(* IEC 61131-3 sources: IRIS-Project/LASAL CONTROL SOFTWARE/LasalProject_2025_09_25/Network, 1 file *)

(* ---- ConfigObjects.st ---- *)
FUNCTION GLOBAL TAB TASK_CONF
_K_TASK, _K_REAL,
_K_END_VAR,

_K_TASK, _K_CYCLIC,
_K_END_VAR,

_K_TASK, _K_BACKGROUND,
_K_END_VAR,

_K_END_CONF
END_FUNCTION

FUNCTION GLOBAL TAB IPR_CONF
_K_IPR
	0$UINT,
_K_END_VAR,
_K_END_CONF
END_FUNCTION

FUNCTION GLOBAL TAB CONFIG_TABLES
00114$UINT,
0$UINT, 1, 58, "_AXISBASE",
0$UINT, 0, 4, "_CAN",
0$UINT, 1, 10, "_CANLIB",
0$UINT, 1, 0, "_CHECKSUM",
0$UINT, 1, 20, "_FILESYS",
0$UINT, 0, 5, "_LINKER",
0$UINT, 1, 0, "_LMCABSENCODER",
0$UINT, 1, 114, "_LMCAXIS",
0$UINT, 2, 105, "_LMCAXISBASE",
0$UINT, 1, 32, "_LMCAXISREF",
0$UINT, 1, 40, "_LMCAXISVIS",
0$UINT, 1, 62, "_LMCAXISVISINT",
0$UINT, 1, 0, "_LMCAXISVISLOGHANDLE",
0$UINT, 1, 0, "_LMCAXISVISLOGVIEWER",
0$UINT, 1, 13, "_LMCAXISVISPARA",
0$UINT, 1, 1, "_LMCAXISVOVMONITORING",
0$UINT, 1, 75, "_LMCMATHFUNCTIONS",
0$UINT, 1, 0, "_LMCMODULEBASE",
0$UINT, 1, 0, "_LMCPUBLISHER",
0$UINT, 1, 11, "_LMCREFBASE",
0$UINT, 1, 21, "_LMCSAFETY",
0$UINT, 1, 36, "_MODBUSTCPSLAVE",
0$UINT, 1, 1, "_MULTITASK",
0$UINT, 0, 5, "_OSKERNEL",
0$UINT, 1, 34, "_SERLIB",
0$UINT, 0, 0, "_STDLIB",
0$UINT, 0, 0, "_SYSMSG",
0$UINT, 1, 1, "_TASKOBJECTCONTROL",
0$UINT, 1, 38, "_TCPIP_SERVER",
0$UINT, 1, 18, "AI084",
0$UINT, 1, 21, "ASCII_BIN",
0$UINT, 0, 0, "ATTUATORE",
0$UINT, 0, 0, "AUTOMANSELECTOR",
0$UINT, 0, 0, "AUTOMATIC_STEP_SETTINGS",
0$UINT, 2, 1, "BUSINTERFACESDIASINTERNAL",
0$UINT, 1, 46, "CONTROLLER",
0$UINT, 0, 0, "CONTROLLOSERVERMODBUS",
0$UINT, 1, 1, "CP112_IOS",
0$UINT, 0, 4, "CRITICALSECTION",
0$UINT, 1, 12, "DI160",
0$UINT, 2, 33, "DIASMASTER",
0$UINT, 1, 83, "DIASMASTERC",
0$UINT, 2, 25, "DIASMASTERMAIN",
0$UINT, 1, 0, "DIASMASTERPOSTSCAN",
0$UINT, 0, 0, "DISCHARGETIMER",
0$UINT, 1, 11, "EEPROM",
0$UINT, 0, 0, "ESTOPMANAGER",
0$UINT, 0, 0, "EXACTSTEP",
0$UINT, 0, 0, "HOLDINGREGISTER",
0$UINT, 0, 0, "HOLDINGREGISTER_2",
0$UINT, 0, 0, "HOLDINGREGISTER_3",
0$UINT, 1, 21, "HUB_BASE",
0$UINT, 2, 11, "HUB_BASE_ROOT",
0$UINT, 2, 36, "HWBASE",
0$UINT, 2, 56, "HWBASECDIAS",
0$UINT, 1, 0, "HWCLOGGING",
0$UINT, 5, 21, "HWCONTROL",
0$UINT, 1, 10, "HWCONTROLBASE",
0$UINT, 1, 0, "HWRTPOSTSCAN",
0$UINT, 1, 6, "I2CCDIAS",
0$UINT, 0, 0, "INPUTREGISTER",
0$UINT, 0, 0, "IRRADIATIONMANAGER",
0$UINT, 1, 0, "LOGIC_NOT",
0$UINT, 1, 0, "LOGIC_XOR",
0$UINT, 0, 0, "MAINSEQUENCE",
0$UINT, 0, 0, "MANAGER_GLOBALE",
0$UINT, 0, 0, "MANAGER_MANUAL_MOTOR",
0$UINT, 0, 0, "MANAGERMOTORI",
0$UINT, 0, 0, "MANUAL_MOTOR",
0$UINT, 0, 0, "MANUAL_MOTORBT",
0$UINT, 0, 0, "MANUAL_STEP_SETTINGS",
0$UINT, 0, 0, "MANUALMOTOR_CBCM",
0$UINT, 0, 0, "MANUALMOTOR_DB",
0$UINT, 1, 22, "MERKEREX",
0$UINT, 0, 0, "MODE_SELECTOR_CLASS",
0$UINT, 0, 0, "MOTORE_M1",
0$UINT, 0, 0, "MOTORE_M2",
0$UINT, 0, 0, "MOTORE_M3",
0$UINT, 0, 0, "MOTORE_M4",
0$UINT, 0, 0, "MOTORE_M5",
0$UINT, 0, 0, "MOTORE_M6",
0$UINT, 0, 0, "MOTORE_M7",
0$UINT, 0, 0, "MOVETIMER",
0$UINT, 0, 0, "MPS",
0$UINT, 0, 0, "RACK12V",
0$UINT, 1, 9, "RAMFILE",
0$UINT, 0, 0, "RESET",
0$UINT, 3, 19, "SAFETYCDIAS_BASE",
0$UINT, 2, 26, "SAFETYMANAGER",
0$UINT, 1, 4, "SAFETYUDP",
0$UINT, 1, 60, "SDIASBASE",
0$UINT, 1, 10, "SDIASHUBBASE",
0$UINT, 1, 97, "SDIASMANAGER",
0$UINT, 2, 6, "SDIASPLC",
0$UINT, 0, 42, "SIGCLIB",
0$UINT, 1, 6, "ST151",
0$UINT, 1, 0, "ST151_INTVISU",
0$UINT, 1, 4, "ST151BASE",
0$UINT, 1, 3, "STEPPERCONTROL",
0$UINT, 1, 11, "STRING",
0$UINT, 1, 85, "STRINGINTERNAL",
0$UINT, 1, 21, "SYNCCALL",
0$UINT, 1, 5, "SYSDATETIME",
0$UINT, 0, 1, "SYSTEM",
0$UINT, 1, 1, "TIMEDATELIB",
0$UINT, 1, 0, "TIMERLIB",
0$UINT, 1, 44, "TO127",
0$UINT, 2, 20, "VARAN_BASE",
0$UINT, 3, 7, "VARANMANAGER",
0$UINT, 2, 7, "VARANMANAGER_1",
0$UINT, 1, 26, "VARANMANAGER_BASE",
0$UINT, 1, 3, "VIRTUALBASEINIT",
0$UINT, 2, 11, "WATCHDOGDIAS",
0$UINT, 1, 1, "XXXBASE_IOS",
ONE_CFG$UINT, 0, 0, "ONE_Comunicazione_ModBus",
ONE_CFG$UINT, 0, 0, "ONE_HW_Network",
ONE_CFG$UINT, 0, 0, "ONE_IRIS_MANAGER",
ONE_CFG$UINT, 0, 0, "ONE_Manual",
ONE_CFG$UINT, 0, 0, "ONE_Profili_Assi",
ONE_CFG$UINT, 0, 0, "ONE_Settings",
ONE_CFG$UINT, 0, 0, "ONE_Timer",
TASK_CFG$UINT, 0, 0, "TASK_CONF",
IPR_CFG$UINT, 0, 0, "IPR_CONF",
PRJ_CFG$UINT, 0, 0, "v1",
END_FUNCTION

#ifdef __LSLLDR_IOELEMENTS__
FUNCTION GLOBAL TAB _IO_ELEMENTS_TAB
0001$UINT, 0133$UINT,
"**IOCONN_EMPTY**", "ST1517.Input1",
"IO_Element", "_LMCAxis_M1.Control",
"IO_Element0", "ST1511.AxError",
"IO_Element1", "ST1511.Enable",
"IO_Element10", "_LMCAxis_M7.Control",
"IO_Element100", "_LMCAxis_M6.ActPos",
"IO_Element101", "Manager_globale1.enable",
"IO_Element102", "_LMCAxis_M1.ActPos",
"IO_Element103", "_LMCAxis_M2.ActPos",
"IO_Element104", "_LMCAxis_M3.ActPos",
"IO_Element105", "_LMCAxis_M4.ActPos",
"IO_Element106", "_LMCAxis_M5.ActPos",
"IO_Element107", "_LMCAxis_M6.ActPos",
"IO_Element108", "_LMCAxis_M7.ActPos",
"IO_Element109", "TO1271.Output4",
"IO_Element11", "ST1511.ActPosition",
"IO_Element110", "TO1271.Output8",
"IO_Element111", "TO1271.Output11",
"IO_Element112", "TO1271.Output10",
"IO_Element113", "ST1516.MaxCurrent",
"IO_Element114", "MPS1.ReqToMPS",
"IO_Element115", "Motore_M51.s_TabletTimer",
"IO_Element116", "Manager_globale1.ComandoIrradiation",
"IO_Element117", "MoveTimer1.s_StartStopTimer",
"IO_Element118", "MoveTimer1.s_StartStopTimer",
"IO_Element119", "MainSequence1.s_EasyGUI",
"IO_Element12", "_LMCAxis_M1.Control",
"IO_Element120", "IrradiationTimers.s_EasyGUI",
"IO_Element121", "Reset1.s_ResetT",
"IO_Element122", "IrradiationTimers.s_TimerStartStop",
"IO_Element123", "ST1514.MaxCurrent",
"IO_Element124", "ST1511.MaxCurrent",
"IO_Element125", "ST1513.MaxCurrent",
"IO_Element126", "ST1516.MaxCurrent",
"IO_Element127", "ST1515.MaxCurrent",
"IO_Element128", "ST1512.MaxCurrent",
"IO_Element129", "MoveTimer1.s_1_3_pelletMode",
"IO_Element13", "ST1511.Input2",
"IO_Element130", "IrradiationTimers.s_1_3_pelletMode",
"IO_Element14", "Motore_M11.M1_Correction_Step",
"IO_Element15", "ST1512.ActPosition",
"IO_Element16", "ST1511.Input1",
"IO_Element17", "ST1511.Input2",
"IO_Element18", "Motore_M41.M4_Correction_Step",
"IO_Element19", "DI1601.Input3",
"IO_Element2", "ST1511.SetFreqOut",
"IO_Element20", "ST1512.AxError",
"IO_Element21", "ST1512.Enable",
"IO_Element22", "ST1512.SetFreqOut",
"IO_Element23", "ST1512.ErrorQuit",
"IO_Element24", "ST1513.ActPosition",
"IO_Element25", "ST1513.AxError",
"IO_Element26", "ST1513.Enable",
"IO_Element27", "ST1513.SetFreqOut",
"IO_Element28", "ST1513.ErrorQuit",
"IO_Element29", "ST1514.ActPosition",
"IO_Element3", "ST1511.ErrorQuit",
"IO_Element30", "ST1514.AxError",
"IO_Element31", "ST1514.Enable",
"IO_Element32", "ST1514.SetFreqOut",
"IO_Element33", "ST1514.ErrorQuit",
"IO_Element34", "ST1512.Input2",
"IO_Element35", "TO1271.Output2",
"IO_Element36", "ST1513.Input1",
"IO_Element37", "ST1513.Input2",
"IO_Element38", "ST1514.Input1",
"IO_Element39", "TO1271.Output3",
"IO_Element4", "_LMCAxis_M2.Control",
"IO_Element40", "TO1271.Output1",
"IO_Element41", "TO1271.Output5",
"IO_Element42", "TO1271.Output6",
"IO_Element43", "TO1271.Output7",
"IO_Element44", "ST1515.ActPosition",
"IO_Element45", "ST1515.AxError",
"IO_Element46", "ST1515.Enable",
"IO_Element47", "ST1515.SetFreqOut",
"IO_Element48", "ST1515.ErrorQuit",
"IO_Element49", "ST1515.Input1",
"IO_Element5", "_LMCAxis_M3.Control",
"IO_Element50", "ST1516.Input1",
"IO_Element51", "ST1516.Input2",
"IO_Element52", "ST1513.MaxCurrent",
"IO_Element53", "ST1516.ActPosition",
"IO_Element54", "ST1516.AxError",
"IO_Element55", "ST1516.Enable",
"IO_Element56", "ST1516.SetFreqOut",
"IO_Element57", "ST1516.ErrorQuit",
"IO_Element58", "ST1511.MaxCurrent",
"IO_Element59", "ST1515.MaxCurrent",
"IO_Element6", "_LMCAxis_M4.Control",
"IO_Element60", "_LMCAxis_M5.ActPos",
"IO_Element61", "_LMCAxis_M1.ActPos",
"IO_Element62", "_LMCAxis_M3.ActPos",
"IO_Element63", "ST1517.ActPosition",
"IO_Element64", "ST1517.AxError",
"IO_Element65", "ST1517.Enable",
"IO_Element66", "ST1517.SetFreqOut",
"IO_Element67", "ST1517.ErrorQuit",
"IO_Element68", "ST1517.Input1",
"IO_Element69", "ST1517.Input2",
"IO_Element7", "_LMCAxis_M5.Control",
"IO_Element70", "_LMCAxis_M7.ActPos",
"IO_Element71", "ST1514.MaxCurrent",
"IO_Element72", "Motore_M31.M3_Correction_Step",
"IO_Element73", "Motore_M51.M5_ChargingCorrection_step_1",
"IO_Element74", "Motore_M51.M5_ChargingCorrection_step_2",
"IO_Element75", "Motore_M51.M5_ChargingCorrection_step_3",
"IO_Element76", "Motore_M51.M5_IrradiationCorrection_step_1",
"IO_Element77", "Motore_M51.M5_IrradiationCorrection_step_2",
"IO_Element78", "_LMCAxis_M2.Control",
"IO_Element79", "Motore_M51.M5_IrradiationCorrection_step_3",
"IO_Element8", "_LMCAxis_M6.Control",
"IO_Element80", "Motore_M51.M5_DischargeCorrection_step",
"IO_Element81", "ST1512.Input2",
"IO_Element82", "_LMCAxis_M3.Control",
"IO_Element83", "_LMCAxis_M4.Control",
"IO_Element84", "DI1601.Input1",
"IO_Element85", "TO1271.Output9",
"IO_Element86", "_LMCAxis_M5.Control",
"IO_Element87", "_LMCAxis_M6.Control",
"IO_Element88", "_LMCAxis_M7.Control",
"IO_Element89", "ST1513.Input1",
"IO_Element9", "ST1511.Input1",
"IO_Element90", "ST1513.Input2",
"IO_Element91", "ST1514.Input1",
"IO_Element92", "ST1515.Input1",
"IO_Element93", "ST1516.Input1",
"IO_Element94", "ST1516.Input2",
"IO_Element95", "Motore_M51.s_tablet_irradiation_position",
"IO_Element96", "DischargeTimer1.s_StartStopTimer",
"IO_Element97", "_LMCAxis_M2.ActPos",
"IO_Element98", "ManagerMotori1.From_MPS",
"IO_Element99", "_LMCAxis_M4.ActPos",
0134$UINT,
"**IOCONN_EMPTY**", "M7_Target_Block.M_LS_1",
"**IOCONN_EMPTY**", "M7_Target_Block.M_LS_2",
"IO_Element", "Motore_M11.Comando_M1",
"IO_Element0", "StepperControl_M1.HWErrors",
"IO_Element1", "StepperControl_M1.Active",
"IO_Element10", "Motore_M71.Comando_M7",
"IO_Element100", "Motore_M61.SetPosition_Controller",
"IO_Element101", "AutoManSelector1.toAutomatic",
"IO_Element102", "M1_Charge_Slider.setPositionController",
"IO_Element103", "M2_Charge_Buffer.setPositionController",
"IO_Element104", "M3_Discharge_Slider.setPositionController",
"IO_Element105", "M4_Discharge_Buffer.setPositionController",
"IO_Element106", "M5_Central_Movement.setPositionController",
"IO_Element107", "M6_Longitudinal_axis.setPositionController",
"IO_Element108", "M7_Target_Block.setPositionController",
"IO_Element109", "Rack12V1.ToPLC",
"IO_Element11", "_LMCAxis_M1.ActPosition",
"IO_Element110", "ManagerMotori1.LED_Rosso",
"IO_Element111", "ManagerMotori1.LED_Arancione",
"IO_Element112", "ManagerMotori1.LED_Verde",
"IO_Element113", "MPS1.To_CameraAlignment_Power",
"IO_Element114", "ManagerMotori1.c_MPS_Req",
"IO_Element115", "IrradiationTimers.NrIrrTablets",
"IO_Element116", "IrradiationTimers.SetStartStopIrr",
"IO_Element117", "Motore_M51.c_TimerMov",
"IO_Element118", "Motore_M41.c_TimerMov",
"IO_Element119", "AutoManSelector1.c_EasyGUIEn_MainS",
"IO_Element12", "M1_Charge_Slider.Comando_Motore",
"IO_Element120", "AutoManSelector1.c_EasyGUIEn_IrrT",
"IO_Element121", "Manager_globale1.c_ResetTimer",
"IO_Element122", "Motore_M51.c_TimerIrr",
"IO_Element123", "M4_Discharge_Buffer.c_MaxCurrent",
"IO_Element124", "M1_Charge_Slider.c_MaxCurrent",
"IO_Element125", "M3_Discharge_Slider.c_MaxCurrent",
"IO_Element126", "M6_Longitudinal_axis.c_MaxCurrent",
"IO_Element127", "M5_Central_Movement.c_MaxCurrent",
"IO_Element128", "M2_Charge_Buffer.c_MaxCurrent",
"IO_Element129", "ManagerMotori1.c_1_3_pelletMode_TimerMov",
"IO_Element13", "Motore_M11.M1_LS_2",
"IO_Element130", "ManagerMotori1.c_1_3_pelletMode_TimerIrr",
"IO_Element14", "Automatic_Step_Settings1.c_M1_Correction_Step",
"IO_Element15", "_LMCAxis_M2.ActPosition",
"IO_Element16", "M1_Charge_Slider.M_LS_1",
"IO_Element17", "M1_Charge_Slider.M_LS_2",
"IO_Element18", "Automatic_Step_Settings1.c_M4_Correction_Step",
"IO_Element19", "Manager_globale1.Reset_IN",
"IO_Element2", "StepperControl_M1.OutputSignal",
"IO_Element20", "StepperControl_M2.HWErrors",
"IO_Element21", "StepperControl_M2.Active",
"IO_Element22", "StepperControl_M2.OutputSignal",
"IO_Element23", "StepperControl_M2.HWErrorQuit",
"IO_Element24", "_LMCAxis_M3.ActPosition",
"IO_Element25", "StepperControl_M3.HWErrors",
"IO_Element26", "StepperControl_M3.Active",
"IO_Element27", "StepperControl_M3.OutputSignal",
"IO_Element28", "StepperControl_M3.HWErrorQuit",
"IO_Element29", "_LMCAxis_M4.ActPosition",
"IO_Element3", "StepperControl_M1.HWErrorQuit",
"IO_Element30", "StepperControl_M4.HWErrors",
"IO_Element31", "StepperControl_M4.Active",
"IO_Element32", "StepperControl_M4.OutputSignal",
"IO_Element33", "StepperControl_M4.HWErrorQuit",
"IO_Element34", "Motore_M21.M2_LS",
"IO_Element35", "Attuatore1.R_aus_1",
"IO_Element36", "Motore_M31.M3_LS_1",
"IO_Element37", "Motore_M31.M3_LS_2",
"IO_Element38", "Motore_M41.M4_LS",
"IO_Element39", "Attuatore1.R_aus_2",
"IO_Element4", "Motore_M21.Comando_M2",
"IO_Element40", "Attuatore1.R_p",
"IO_Element41", "Attuatore2.R_p",
"IO_Element42", "Attuatore2.R_aus_1",
"IO_Element43", "Attuatore2.R_aus_2",
"IO_Element44", "_LMCAxis_M5.ActPosition",
"IO_Element45", "StepperControl_M5.HWErrors",
"IO_Element46", "StepperControl_M5.Active",
"IO_Element47", "StepperControl_M5.OutputSignal",
"IO_Element48", "StepperControl_M5.HWErrorQuit",
"IO_Element49", "Motore_M51.M5_LS",
"IO_Element5", "Motore_M31.Comando_M3",
"IO_Element50", "Motore_M61.M6_LS_1",
"IO_Element51", "Motore_M61.M6_LS_2",
"IO_Element52", "Motore_M31.c_MaxCurrent",
"IO_Element53", "_LMCAxis_M6.ActPosition",
"IO_Element54", "StepperControl_M6.HWErrors",
"IO_Element55", "StepperControl_M6.Active",
"IO_Element56", "StepperControl_M6.OutputSignal",
"IO_Element57", "StepperControl_M6.HWErrorQuit",
"IO_Element58", "Motore_M11.c_MaxCurrent",
"IO_Element59", "Motore_M51.c_MaxCurrent",
"IO_Element6", "Motore_M41.Comando_M4",
"IO_Element60", "Motore_M51.SetPosition_Controller",
"IO_Element61", "Motore_M11.SetPosition_Controller",
"IO_Element62", "Motore_M31.SetPositionController",
"IO_Element63", "_LMCAxis_M7.ActPosition",
"IO_Element64", "StepperControl_M7.HWErrors",
"IO_Element65", "StepperControl_M7.Active",
"IO_Element66", "StepperControl_M7.OutputSignal",
"IO_Element67", "StepperControl_M7.HWErrorQuit",
"IO_Element68", "Motore_M71.M7_LS_1",
"IO_Element69", "Motore_M71.M7_LS_2",
"IO_Element7", "Motore_M51.Comando_M5",
"IO_Element70", "Motore_M71.SetPositionController",
"IO_Element71", "Motore_M41.c_MaxCurrent",
"IO_Element72", "Automatic_Step_Settings1.c_M3_Correction_Step",
"IO_Element73", "Automatic_Step_Settings1.c_M5_ChargingCorrection_Step_1",
"IO_Element74", "Automatic_Step_Settings1.c_M5_ChargingCorrection_Step_2",
"IO_Element75", "Automatic_Step_Settings1.c_M5_ChargingCorrection_Step_3",
"IO_Element76", "Automatic_Step_Settings1.c_M5_IrradiationCorrection_Step_1",
"IO_Element77", "Automatic_Step_Settings1.c_M5_IrradiationCorrection_Step_2",
"IO_Element78", "M2_Charge_Buffer.Comando_Motore",
"IO_Element79", "Automatic_Step_Settings1.c_M5_IrradiationCorrection_step_3",
"IO_Element8", "Motore_M61.Comando_M6",
"IO_Element80", "Automatic_Step_Settings1.c_M5_DischargingCorrection_step",
"IO_Element81", "M2_Charge_Buffer.M_LS",
"IO_Element82", "M3_Discharge_Slider.Comando_Motore",
"IO_Element83", "M4_Discharge_Buffer.Comando_Motore",
"IO_Element84", "MPS1.ACKFromMPS",
"IO_Element85", "MPS1.c_ReqToMPS",
"IO_Element86", "M5_Central_Movement.Comando_Motore",
"IO_Element87", "M6_Longitudinal_axis.Comando_Motore",
"IO_Element88", "M7_Target_Block.Comando_Motore",
"IO_Element89", "M3_Discharge_Slider.M_LS_2",
"IO_Element9", "Motore_M11.M1_LS_1",
"IO_Element90", "M3_Discharge_Slider.M_LS_1",
"IO_Element91", "M4_Discharge_Buffer.M_LS",
"IO_Element92", "M5_Central_Movement.M_LS",
"IO_Element93", "M6_Longitudinal_axis.M_LS_1",
"IO_Element94", "M6_Longitudinal_axis.M_LS_2",
"IO_Element95", "IrradiationTimers.TabletInIrrPos",
"IO_Element96", "Motore_M41.c_TimerDis",
"IO_Element97", "Motore_M21.SetPosition_Controller",
"IO_Element98", "MPS1.To_Manager_Motori",
"IO_Element99", "Motore_M41.SetPositionController",
END_FUNCTION
#endif //__LSLLDR_IOELEMENTS__

FUNCTION GLOBAL TAB CH_REDIRECT_EMB_TAB
0000$UINT,
00012$UINT,
"_TCPIP_SERVER;SEMANAME01", "\STRSEMANAME01.DATA",
"_TCPIP_SERVER;SEMANAME02", "\STRSEMANAME02.DATA",
"_TCPIP_SERVER;TASKNAME", "\STRTASKNAME.DATA",
"AI084;SERIALNO", "\SERIALNOSTR.DATA",
"DI160;SERIALNO", "\SERIALNOSTR.DATA",
"HWBASECDIAS;SERIALNO", "\SERIALNOSTR.DATA",
"SAFETYCDIAS_BASE;SERIALNO", "\SERIALNOSTR.DATA",
"SDIASBASE;SERIALNO", "\SERIALNOSTR.DATA",
"ST151;SERIALNO", "\SERIALNOSTR.DATA",
"ST151BASE;SERIALNO", "\SERIALNOSTR.DATA",
"TO127;SERIALNO", "\SERIALNOSTR.DATA",
"VARAN_BASE;SERIALNO", "\SERIALNOSTR.DATA",
END_FUNCTION
